(* IEC 61131-3 sources: codesys-framework/txt/application/WeVe Core (library)/30 Module/FB_Module/State, 9 files *)

(* ---- ProcessDisable.method.st ---- *)
METHOD PROTECTED ProcessDisable
VAR_INPUT
END_VAR

// --- BEGIN IMPLEMENTATION ---

_xEnabled := FALSE;
_eState := E_ModuleStates.Idle;

(* ---- ProcessEnable.method.st ---- *)
METHOD PROTECTED ProcessEnable
VAR_INPUT
END_VAR

// --- BEGIN IMPLEMENTATION ---

_xEnabled := TRUE;
_eState := E_ModuleStates.Standby;

(* ---- ProcessExecute.method.st ---- *)
METHOD PROTECTED ProcessExecute
VAR_INPUT
END_VAR

// --- BEGIN IMPLEMENTATION ---

// Commando klaar, gefaald, afgebroken of timeout: terug naar Standby
IF _fbCmd.Active = 0 THEN
	_xBusy := FALSE;
	_eState := E_ModuleStates.Standby;
	RETURN;
END_IF

_xBusy := TRUE;
ExecuteCommand(iCmd := _fbCmd.Active);

(* ---- ProcessIdle.method.st ---- *)
METHOD PROTECTED ProcessIdle
VAR_INPUT
END_VAR

// --- BEGIN IMPLEMENTATION ---

;

(* ---- ProcessQuickStop.method.st ---- *)
METHOD Protected ProcessQuickStop
VAR_INPUT
END_VAR

// --- BEGIN IMPLEMENTATION ---

// QuickStop is dominant: het actieve commando wordt afgebroken (Aborted).
// Een afgeleide module die hier overschrijft, zet zelf haar uitgangen veilig en roept SUPER^.ProcessQuickStop() aan.
_fbCmd.Abort();

_eState := E_ModuleStates.Invalid;

(* ---- ProcessReset.method.st ---- *)
METHOD PROTECTED ProcessReset
VAR_INPUT
END_VAR

// --- BEGIN IMPLEMENTATION ---

_eState := E_ModuleStates.Initialize;

(* ---- ProcessStandby.method.st ---- *)
METHOD PROTECTED ProcessStandby
VAR_INPUT
END_VAR

// --- BEGIN IMPLEMENTATION ---

_xDone := FALSE;
_xBusy := FALSE;

(* ---- ProcessState.method.st ---- *)
METHOD PRIVATE ProcessState
VAR_INPUT
END_VAR

// --- BEGIN IMPLEMENTATION ---

CASE _eState OF

	E_ModuleStates.Invalid 			: ;
	E_ModuleStates.Initialize 		: ;
	E_ModuleStates.Idle 			: ProcessIdle();
	E_ModuleStates.Enable 			: ProcessEnable();
	E_ModuleStates.Standby 			: ProcessStandby();
	E_ModuleStates.Execute 			: ProcessExecute();
	E_ModuleStates.Disable 			: ProcessDisable();
	E_ModuleStates.Stop 			: ProcessStop();
	E_ModuleStates.QuickStop 		: ProcessQuickStop();
	E_ModuleStates.Reset 			: ProcessReset();

END_CASE

(* ---- ProcessStop.method.st ---- *)
METHOD PROTECTED ProcessStop
VAR_INPUT
END_VAR

// --- BEGIN IMPLEMENTATION ---

// Stop is dominant: het actieve commando wordt afgebroken (Aborted).
// Een afgeleide module die hier overschrijft, zet zelf haar uitgangen veilig en roept SUPER^.ProcessStop() aan.
_fbCmd.Abort();

_eState := E_ModuleStates.Disable;
